(* IEC 61131-3 sources: llm-plc-st-eval/data/processed_definitivo/qwen2.5-coder_14b/I8/few_shot, 3 files *)

(* ---- ejec_1.st ---- *)
FUNCTION_BLOCK FB_Compresor
VAR_INPUT
    pOilOk : BOOL; (* Presión de aceite correcta *)
    tempOk : BOOL; (* Temperatura correcta *)
    sinAlm : BOOL; (* Ausencia de alarmas *)
    btnMarcha : BOOL; (* Botón de marcha *)
    btnParo : BOOL; (* Botón de paro *)
END_VAR
VAR_OUTPUT
    comp : BOOL; (* Compresor *)
    causaBloqueo : INT; (* Causa de bloqueo *)
END_VAR
VAR
    tOilOk : TP; (* Temporizador para presión de aceite *)
    marchaAnt : BOOL; (* Estado anterior del botón de marcha *)
    permisivoOk : BOOL; (* Permiso para arranque *)
END_VAR

(* Temporizador para la presión de aceite *)
tOilOk(IN := pOilOk, PT := T#3S);

(* Determinar si todos los permisivos están cumplidos *)
permisivoOk := tOilOk.Q AND tempOk AND sinAlm;

(* Determinar la causa de bloqueo *)
IF NOT pOilOk THEN
    causaBloqueo := 1;
ELSIF NOT tempOk THEN
    causaBloqueo := 2;
ELSIF NOT sinAlm THEN
    causaBloqueo := 3;
ELSE
    causaBloqueo := 0;
END_IF;

(* Control de arranque y paro del compresor *)
IF btnParo THEN
    comp := FALSE;
ELSIF btnMarcha AND NOT marchaAnt AND permisivoOk THEN
    comp := TRUE;
END_IF;

(* Guardar el estado anterior del botón de marcha *)
marchaAnt := btnMarcha;
END_FUNCTION_BLOCK

(* ---- ejec_2.st ---- *)
FUNCTION_BLOCK FB_Compresor
VAR_INPUT
    pOilOk : BOOL; (* Presión de aceite correcta *)
    tempOk : BOOL; (* Temperatura correcta *)
    sinAlm : BOOL; (* Ausencia de alarmas *)
    btnMarcha : BOOL; (* Botón de marcha *)
    btnParo : BOOL; (* Botón de paro *)
END_VAR
VAR_OUTPUT
    comp : BOOL; (* Compresor *)
    causaBloqueo : INT; (* Causa de bloqueo *)
END_VAR
VAR
    tPresion : TP; (* Temporizador para presión de aceite *)
    marchaAnterior : BOOL; (* Estado anterior del botón de marcha *)
    permisivoCumplido : BOOL; (* Indica si todos los permisivos están cumplidos *)
END_VAR

(* Temporizador para la presión de aceite *)
tPresion(IN := pOilOk, PT := T#3S);

(* Comprobar si todos los permisivos están cumplidos *)
permisivoCumplido := tPresion.Q AND tempOk AND sinAlm;

(* Determinar la causa de bloqueo *)
IF NOT pOilOk THEN
    causaBloqueo := 1;
ELSIF NOT tempOk THEN
    causaBloqueo := 2;
ELSIF NOT sinAlm THEN
    causaBloqueo := 3;
ELSE
    causaBloqueo := 0;
END_IF;

(* Control de arranque y paro del compresor *)
IF btnParo THEN
    comp := FALSE;
ELSIF btnMarcha AND NOT marchaAnterior AND permisivoCumplido THEN
    comp := TRUE;
END_IF;

(* Actualizar el estado anterior del botón de marcha *)
marchaAnterior := btnMarcha;
END_FUNCTION_BLOCK

(* ---- ejec_3.st ---- *)
FUNCTION_BLOCK FB_Compresor
VAR_INPUT
    pOilOk : BOOL; (* Presión de aceite correcta *)
    tempOk : BOOL; (* Temperatura correcta *)
    sinAlm : BOOL; (* Ausencia de alarmas *)
    btnMarcha : BOOL; (* Botón de marcha *)
    btnParo : BOOL; (* Botón de paro *)
END_VAR
VAR_OUTPUT
    comp : BOOL; (* Compresor *)
    causaBloqueo : INT; (* Causa de bloqueo *)
END_VAR
VAR
    tPresion : TP; (* Temporizador para presión de aceite *)
    marchaAnterior : BOOL; (* Estado anterior del botón de marcha *)
    permisivoCumplido : BOOL; (* Indica si todos los permisivos están cumplidos *)
END_VAR

(* Temporizador para la presión de aceite *)
tPresion(IN := pOilOk, PT := T#3S);

(* Determina si todos los permisivos están cumplidos *)
permisivoCumplido := tPresion.Q AND tempOk AND sinAlm;

(* Determina la causa de bloqueo *)
IF NOT pOilOk THEN
    causaBloqueo := 1;
ELSIF NOT tempOk THEN
    causaBloqueo := 2;
ELSIF NOT sinAlm THEN
    causaBloqueo := 3;
ELSE
    causaBloqueo := 0;
END_IF;

(* Control de arranque y paro del compresor *)
IF btnParo THEN
    comp := FALSE;
ELSIF btnMarcha AND NOT marchaAnterior AND permisivoCumplido THEN
    comp := TRUE;
END_IF;

(* Actualiza el estado anterior del botón de marcha *)
marchaAnterior := btnMarcha;
END_FUNCTION_BLOCK
